(* IEC 61131-3 sources: trust-platform/examples/rust_signal/src/generated, 1 file *)

(* ---- rust_pous.st ---- *)
(* GENERATED by trust-runtime from rust/src/lib.rs - do not edit *)
{attribute 'rust'}
FUNCTION_BLOCK MEDIAN5
VAR_INPUT
    EN : BOOL := TRUE;
    x : REAL;
END_VAR
VAR_OUTPUT
    y : REAL;
    mean : REAL;
END_VAR
VAR
    history : ARRAY[0..4] OF REAL;
    next : INT;
    primed : BOOL;
END_VAR
VAR_OUTPUT
    ENO : BOOL;
END_VAR
END_FUNCTION_BLOCK

(* GENERATED by trust-runtime from rust/src/lib.rs - do not edit *)
{attribute 'rust'}
FUNCTION_BLOCK MODBUS_CRC
VAR_INPUT
    EN : BOOL := TRUE;
    frame : ARRAY[0..31] OF BYTE;
    length : INT;
END_VAR
VAR_OUTPUT
    crc : WORD;
    ok : BOOL;
    ENO : BOOL;
END_VAR
END_FUNCTION_BLOCK
